(* IEC 61131-3 sources: 89152_FlorisHendrix_AfstudeerProject/89152_FlorisHendrix_ExamenProject/Stations/MachineControl/MachineControl/Network/XML_Network, 1 file *)

(* ---- ONE_XML_Network_Table.st ---- *)
#define OBJECTS_CONFIG

//Define part of class FileBaseCsv
#define MAX_STRING_LEN    80
#define LF 	          		16#0A		// LF	- LineFeed
#define CR 		          	16#0D		// CR	- Caridge return
#define SEPARATOR  	    	';'

FUNCTION GLOBAL TAB ONE_XML_Network
-1$UINT, 0$UINT,
0$UINT, 0$UINT,

1$UDINT,
TO_UDINT(3416595442), "FileBaseCsv", 0$UINT, 12$UINT, 1$UINT,

_NO_ATTR, TO_UDINT(3500464540), "FILEBASECSV1",

//Internal connections
0$UDINT,
0$UDINT,
0$UDINT,
0$UDINT,

//Initialization values
0$UDINT,
0$UDINT,

//Symbolic initialization values
0$UDINT,
0$UDINT,

//Initialization of string values
0$UDINT,
0$UDINT,

//Configuration of tasks (RealTime, Cyclic, Background)
0$UDINT,
0$UDINT,

0$UDINT,
0$UDINT,

0$UDINT,
0$UDINT,

//External connections
0$UDINT,
0$UDINT,

//Magic internal connections
0$UDINT,
0$UDINT,

//Configuration of timeslots of tasks (RealTime, Cyclic)
#ifdef __LSLLDR_TIMESLOTS__
0$UDINT,
0$UDINT,

0$UDINT,
0$UDINT,

#endif //__LSLLDR_TIMESLOTS__

//MultiMaster connections
#ifdef __LSLLDR_MULTIMASTER__
0$UDINT,
0$UDINT,
#endif //__LSLLDR_MULTIMASTER__

//Configuration for task ID (RealTime, CyclicTime)
#ifdef __LSLLDR_TASKID__
"\\\\TASKS2  "
0$UDINT,
0$UDINT,

0$UDINT,
0$UDINT,

0$UDINT,
0$UDINT,

#endif //__LSLLDR_TASKID__

END_FUNCTION
